(* IEC 61131-3 sources: plc-vscode/tests/st/test-ready/trust-platform/examples/plcopen_motion_single_axis_benchmarks/status_only/src, 2 files *)

(* ---- Globals.st ---- *)
VAR_GLOBAL
    g_motion_bench_cycles : UDINT;
    g_motion_bench_completed_sequences : UDINT;
    g_motion_bench_last_error : WORD;
    g_motion_bench_power_on : BOOL;
    g_motion_bench_is_homed : BOOL;
    g_motion_bench_last_position : REAL;
    g_motion_bench_last_velocity : REAL;
    g_motion_bench_current_step : UINT;
END_VAR

(* ---- Main.st ---- *)
PROGRAM Main
VAR
    Axis : AXIS_REF;
    Power : MC_Power;
    ReadStatus : MC_ReadStatus;
    ReadAxisInfo : MC_ReadAxisInfo;
    ReadMotionState : MC_ReadMotionState;
    ReadAxisError : MC_ReadAxisError;
    ReadActualPosition : MC_ReadActualPosition;
    ReadActualVelocity : MC_ReadActualVelocity;
    Initialized : BOOL;
END_VAR

IF NOT Initialized THEN
    Axis.AxisId := UDINT#1;
    Axis.InternalIndex := UINT#1;
    g_motion_bench_cycles := UDINT#0;
    g_motion_bench_completed_sequences := UDINT#0;
    g_motion_bench_last_error := WORD#16#0000;
    g_motion_bench_power_on := FALSE;
    g_motion_bench_is_homed := FALSE;
    g_motion_bench_last_position := REAL#0.0;
    g_motion_bench_last_velocity := REAL#0.0;
    g_motion_bench_current_step := UINT#1;
    Initialized := TRUE;
END_IF;

g_motion_bench_cycles := g_motion_bench_cycles + UDINT#1;
Power(Axis := Axis, Enable := TRUE);
ReadStatus(Axis := Axis, Enable := TRUE);
ReadAxisInfo(Axis := Axis, Enable := TRUE);
ReadMotionState(Axis := Axis, Enable := TRUE, Source := MC_SOURCE#mcActualValue);
ReadAxisError(Axis := Axis, Enable := TRUE);
ReadActualPosition(Axis := Axis, Enable := TRUE);
ReadActualVelocity(Axis := Axis, Enable := TRUE);

g_motion_bench_completed_sequences := g_motion_bench_cycles;
g_motion_bench_power_on := Power.Status;
g_motion_bench_is_homed := ReadAxisInfo.IsHomed;
g_motion_bench_last_position := ReadActualPosition.Position;
g_motion_bench_last_velocity := ReadActualVelocity.Velocity;
g_motion_bench_current_step := UINT#1;

IF Power.Error THEN
    g_motion_bench_last_error := Power.ErrorID;
ELSIF ReadStatus.Error THEN
    g_motion_bench_last_error := ReadStatus.ErrorID;
ELSIF ReadAxisInfo.Error THEN
    g_motion_bench_last_error := ReadAxisInfo.ErrorID;
ELSIF ReadMotionState.Error THEN
    g_motion_bench_last_error := ReadMotionState.ErrorID;
ELSIF ReadAxisError.AxisErrorID <> WORD#16#0000 THEN
    g_motion_bench_last_error := ReadAxisError.AxisErrorID;
ELSIF ReadActualPosition.Error THEN
    g_motion_bench_last_error := ReadActualPosition.ErrorID;
ELSIF ReadActualVelocity.Error THEN
    g_motion_bench_last_error := ReadActualVelocity.ErrorID;
ELSE
    g_motion_bench_last_error := WORD#16#0000;
END_IF;
END_PROGRAM
